FUNCTION F_DwordToBitReal : REAL
VAR_INPUT
	dwIn : DWORD;
END_VAR
VAR
	pt : POINTER TO REAL;
END_VAR

pt := ADR(dwIn);
F_DwordToBitReal := pt^;

END_FUNCTION

(* stored: Version 1.1.0.1, ProductVersion 3.1.4024.15
   POU F_DwordToBitReal: Id {0c1c280a-ba77-4e36-9578-76dae4150522}, SpecialFunc None *)
